(* Herbal Oil Seperation Process Controlled by Analog Level Sensors *)

PROGRAM main
  VAR
    Inlet AT %QX0.1 : BOOL; (* Master Inlet Valve for Mixture *)
    WaterOutlet AT %QX0.2 : BOOL; (* Outlet Valve for Separated Water *)
    OilOutlet AT %QX0.3 : BOOL;
    TempSensor AT %IW0 : INT;
    LevelSensor AT %IW1 : INT;
  END_VAR

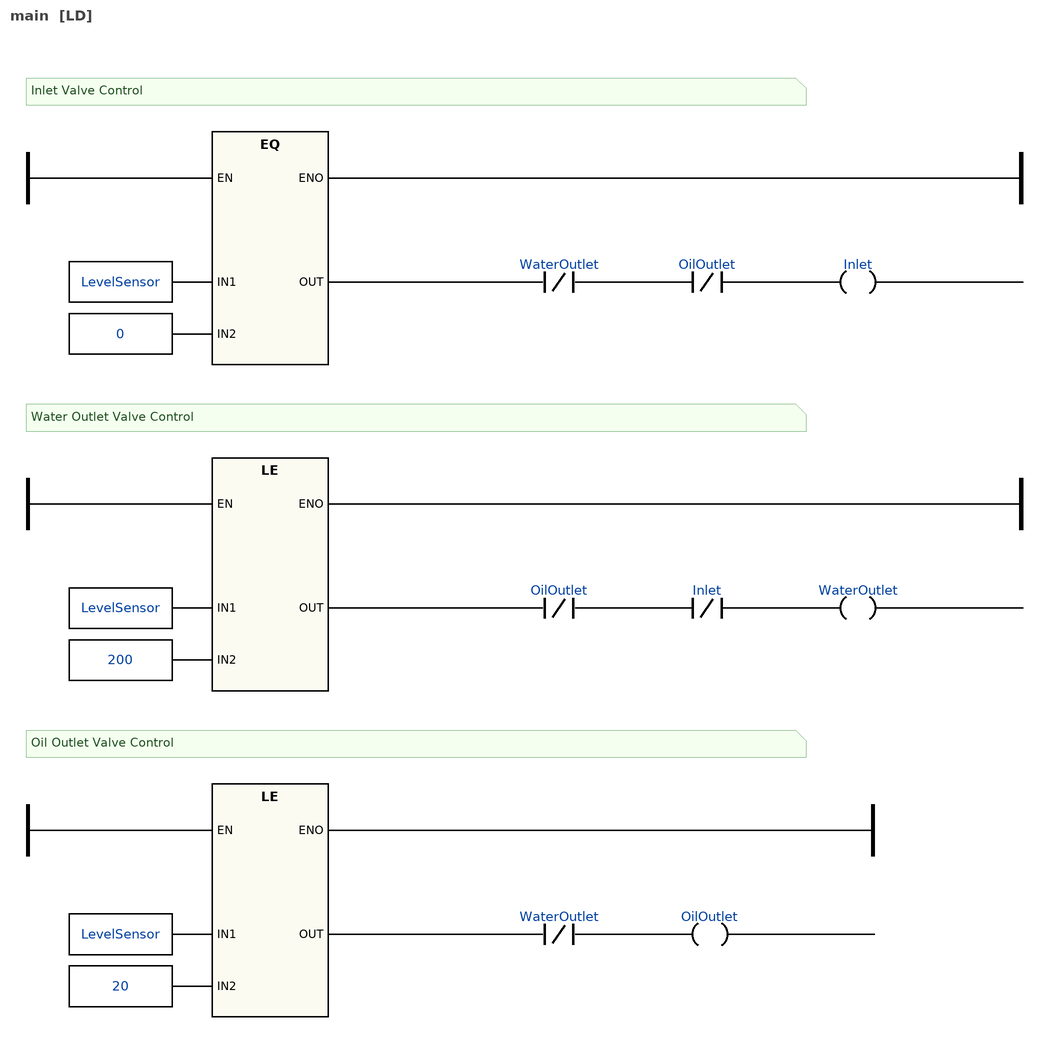
(* LD diagram, written out as Structured Text *)
(* Inlet Valve Control *)
Inlet := LevelSensor = 0 AND NOT WaterOutlet AND NOT OilOutlet;
(* Water Outlet Valve Control *)
WaterOutlet := LevelSensor <= 200 AND NOT OilOutlet AND NOT Inlet;
(* Oil Outlet Valve Control *)
OilOutlet := LevelSensor <= 20 AND NOT WaterOutlet;
END_PROGRAM
